(* LS Electric XG5000 project: KST *)
(* PLC LSPLC *)
(* module base 0 slot 0: 입출력 모듈:KL-5000 (DC 24V 입력 16점/RELAY 출력 12점) *)

PROGRAM NewProgram (* task: 스캔 프로그램 *)
VAR
    Count : INT; (* Source preservation check *)
END_VAR
Count := Count + 1;
END_PROGRAM

PROGRAM AddedST (* task: 스캔 프로그램 *)
VAR
    Count : INT; (* Source preservation check *)
END_VAR
Count := Count + 1;
END_PROGRAM

PROGRAM AddedIL (* task: 스캔 프로그램 *)
VAR
    Count : INT; (* Source preservation check *)
END_VAR
LD Count
ADD 1
ST Count
END_PROGRAM